// TIA Portal V17 export
// export: Created 2026-11-08T05:50:29.3599463Z, ExportSetting WithDefaults, DisplayName Totally Integrated Automation Portal, DisplayVersion V17, DisplayName TIA Portal Openness, DisplayVersion V17, DisplayName TIA Portal Version Control Interface, DisplayVersion V17, DisplayName STEP 7 Professional, DisplayVersion V17, DisplayName STEP 7 Safety, DisplayVersion V17, DisplayName WinCC Professional, DisplayVersion V17
VAR_GLOBAL   // PLC tag table "Pulsadores_y_selectores"
   PB_Marcha AT %M10.0 : Bool;   // Pulsador MARCHA verde (NA)
   PB_Paro AT %M10.1 : Bool;   // Pulsador PARO rojo: 1 = pulsado
END_VAR
